// Worked example: a two-channel emergency stop with contactor feedback, wired the way a
// TwinSAFE project links it, plus the standard PLC signals (Run, ErrAck, Restart).
// The blocks join the group at declaration; call the group before its members.
// CFC twin of PRG_EStopExample: the same wiring as a diagram.
// Toggle the "field" variables online to trial the behaviour and watch the State / Diag outputs.
PROGRAM PRG_EStopExample_CFC
VAR
    // --- simulated field devices (real hardware in a TwinSAFE system)
    eStopChannel1 : BOOL := TRUE; // NC contact, TRUE = not pressed
    eStopChannel2 : BOOL := TRUE;

    // --- standard PLC interface to the TwinSAFE group (linked to standard variables)
    safetyRun : BOOL := TRUE;
    safetyErrAck : BOOL;
    restartButton : BOOL; // 0 -> 1 -> 0 to restart

    // --- TwinSAFE model: the group, then its members (parameters as in the Safety Editor property grid)
    group : T_SafeGroup;
    inputTerminal : T_SafeInputTerminal(group := group); // EL1904
    outputTerminal : T_SafeOutputTerminal(group := group); // EL2904
    eStop : T_SafeEStop(group := group) := (Parameters := (DiscrepancyTime1 := T#500MS, DelayTime := T#1S));

    // --- simulated contactors: pull in 50 ms after the safe output energises; EDM1 = NOT pulled in
    contactorPullIn : TON;
END_VAR

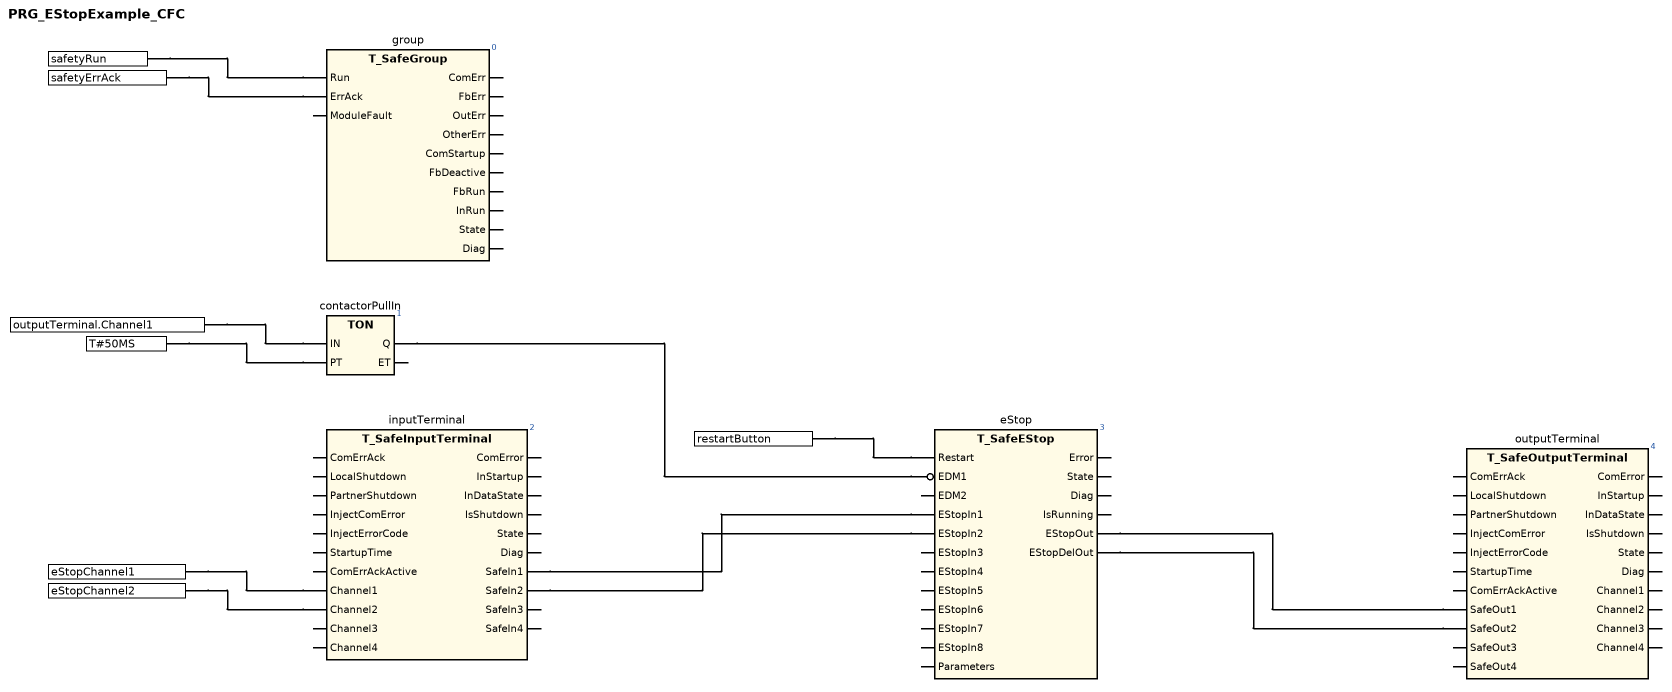
group(Run := safetyRun, ErrAck := safetyErrAck); // T_SafeGroup
contactorPullIn(IN := outputTerminal.Channel1, PT := T#50MS); // TON
inputTerminal(Channel1 := eStopChannel1, Channel2 := eStopChannel2); // T_SafeInputTerminal
eStop(
    Restart := restartButton,
    EDM1 := NOT contactorPullIn.Q,
    EStopIn1 := inputTerminal.SafeIn1,
    EStopIn2 := inputTerminal.SafeIn2); // T_SafeEStop
outputTerminal(SafeOut1 := eStop.EStopOut, SafeOut2 := eStop.EStopDelOut); // T_SafeOutputTerminal

END_PROGRAM

(* stored: Version 1.1.0.1
   POU PRG_EStopExample_CFC: Id {675d26df-9469-584b-b0e9-945da6304417}, SpecialFunc None *)
